// LS Electric XG5000 project: EV_s3
// PLC LSPLC
// module base 0 slot 0: 입출력 모듈:XBC-DR32H (DC 24V 입력, 릴레이 출력 32점)
// module base 0 slot 1: 입력 모듈:XBE-DC16A/B (DC24V 입력, 16점 / DC12/24V 입력, 16점)
// module base 0 slot 2: FEnet:XBL-EMTA (Ethernet 통신 모듈, 전기 Master)
// task INIT: Kind=1 Priority=2

PROGRAM VFD_PARAM (task: 스캔 프로그램)

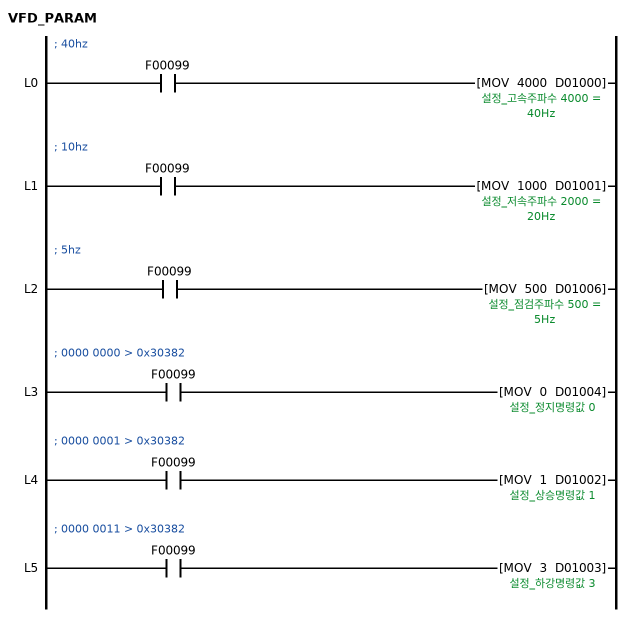
; L0
LOAD      F00099
MOV       4000 D01000	// 설정_고속주파수 4000 = 40Hz
// output comment: 40hz
; L1
LOAD      F00099
MOV       1000 D01001	// 설정_저속주파수 2000 = 20Hz
// output comment: 10hz
; L2
LOAD      F00099
MOV       500 D01006	// 설정_점검주파수 500 = 5Hz
// output comment: 5hz
; L3
LOAD      F00099
MOV       0 D01004	// 설정_정지명령값 0
// output comment: 0000 0000 > 0x30382
; L4
LOAD      F00099
MOV       1 D01002	// 설정_상승명령값 1
// output comment: 0000 0001 > 0x30382
; L5
LOAD      F00099
MOV       3 D01003	// 설정_하강명령값 3
// output comment: 0000 0011 > 0x30382

PROGRAM P00_P_MIRROR (task: 스캔 프로그램)

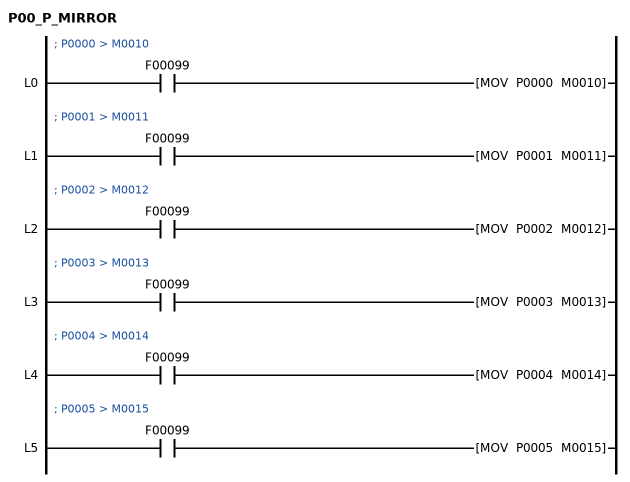
; L0
LOAD      F00099
MOV       P0000 M0010
// output comment: P0000 > M0010
; L1
LOAD      F00099
MOV       P0001 M0011
// output comment: P0001 > M0011
; L2
LOAD      F00099
MOV       P0002 M0012
// output comment: P0002 > M0012
; L3
LOAD      F00099
MOV       P0003 M0013
// output comment: P0003 > M0013
; L4
LOAD      F00099
MOV       P0004 M0014
// output comment: P0004 > M0014
; L5
LOAD      F00099
MOV       P0005 M0015
// output comment: P0005 > M0015

PROGRAM P01_POSITION (task: 스캔 프로그램)

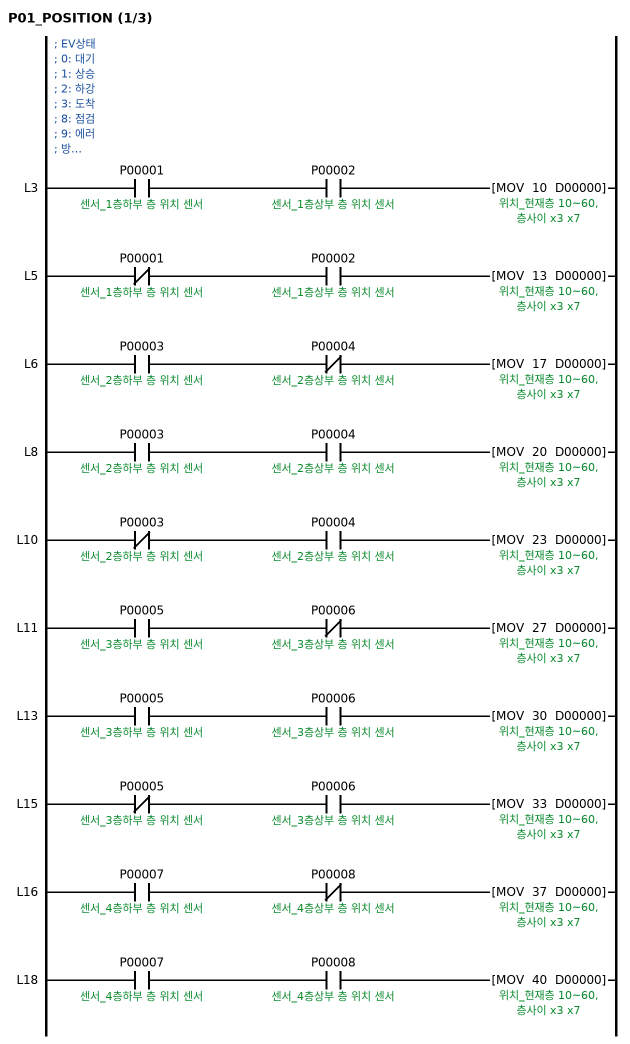
// EV상태
// 0: 대기
// 1: 상승
// 2: 하강
// 3: 도착
// 8: 점검
// 9: 에러
// 방향
// 0: 대기
// 1: 상승
// 2: 하강
// 센서로 인한 현재 위치
; L3
LOAD      P00001	// 센서_1층하부 층 위치 센서
AND       P00002	// 센서_1층상부 층 위치 센서
MOV       10 D00000	// 위치_현재층 10~60, 층사이 x3 x7
; L5
LOAD NOT  P00001	// 센서_1층하부 층 위치 센서
AND       P00002	// 센서_1층상부 층 위치 센서
MOV       13 D00000	// 위치_현재층 10~60, 층사이 x3 x7
; L6
LOAD      P00003	// 센서_2층하부 층 위치 센서
AND NOT   P00004	// 센서_2층상부 층 위치 센서
MOV       17 D00000	// 위치_현재층 10~60, 층사이 x3 x7
; L8
LOAD      P00003	// 센서_2층하부 층 위치 센서
AND       P00004	// 센서_2층상부 층 위치 센서
MOV       20 D00000	// 위치_현재층 10~60, 층사이 x3 x7
; L10
LOAD NOT  P00003	// 센서_2층하부 층 위치 센서
AND       P00004	// 센서_2층상부 층 위치 센서
MOV       23 D00000	// 위치_현재층 10~60, 층사이 x3 x7
; L11
LOAD      P00005	// 센서_3층하부 층 위치 센서
AND NOT   P00006	// 센서_3층상부 층 위치 센서
MOV       27 D00000	// 위치_현재층 10~60, 층사이 x3 x7
; L13
LOAD      P00005	// 센서_3층하부 층 위치 센서
AND       P00006	// 센서_3층상부 층 위치 센서
MOV       30 D00000	// 위치_현재층 10~60, 층사이 x3 x7
; L15
LOAD NOT  P00005	// 센서_3층하부 층 위치 센서
AND       P00006	// 센서_3층상부 층 위치 센서
MOV       33 D00000	// 위치_현재층 10~60, 층사이 x3 x7
; L16
LOAD      P00007	// 센서_4층하부 층 위치 센서
AND NOT   P00008	// 센서_4층상부 층 위치 센서
MOV       37 D00000	// 위치_현재층 10~60, 층사이 x3 x7
; L18
LOAD      P00007	// 센서_4층하부 층 위치 센서
AND       P00008	// 센서_4층상부 층 위치 센서
MOV       40 D00000	// 위치_현재층 10~60, 층사이 x3 x7

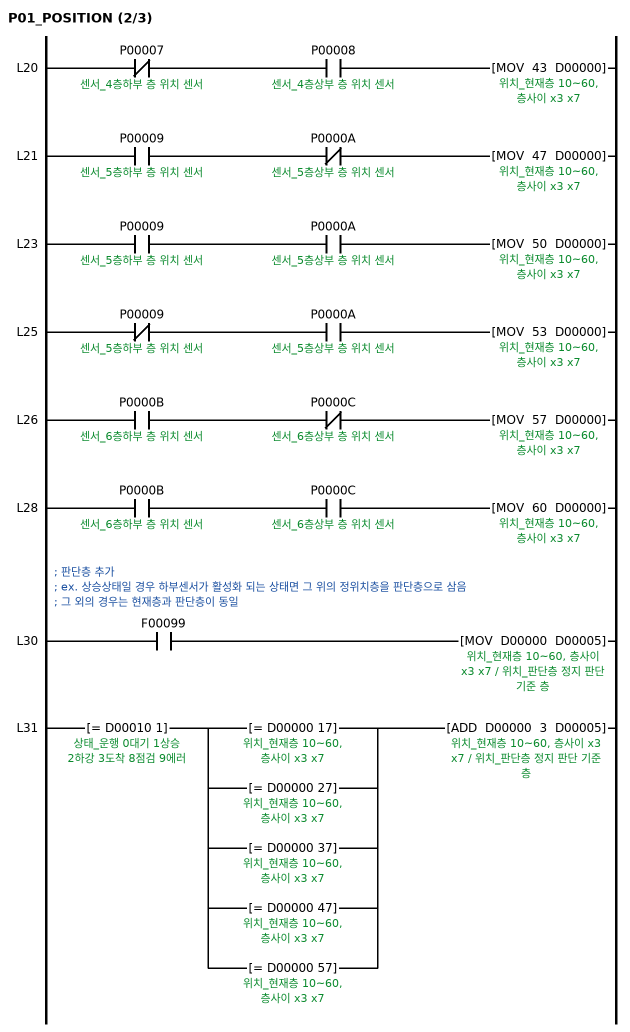
; L20
LOAD NOT  P00007	// 센서_4층하부 층 위치 센서
AND       P00008	// 센서_4층상부 층 위치 센서
MOV       43 D00000	// 위치_현재층 10~60, 층사이 x3 x7
; L21
LOAD      P00009	// 센서_5층하부 층 위치 센서
AND NOT   P0000A	// 센서_5층상부 층 위치 센서
MOV       47 D00000	// 위치_현재층 10~60, 층사이 x3 x7
; L23
LOAD      P00009	// 센서_5층하부 층 위치 센서
AND       P0000A	// 센서_5층상부 층 위치 센서
MOV       50 D00000	// 위치_현재층 10~60, 층사이 x3 x7
; L25
LOAD NOT  P00009	// 센서_5층하부 층 위치 센서
AND       P0000A	// 센서_5층상부 층 위치 센서
MOV       53 D00000	// 위치_현재층 10~60, 층사이 x3 x7
; L26
LOAD      P0000B	// 센서_6층하부 층 위치 센서
AND NOT   P0000C	// 센서_6층상부 층 위치 센서
MOV       57 D00000	// 위치_현재층 10~60, 층사이 x3 x7
; L28
LOAD      P0000B	// 센서_6층하부 층 위치 센서
AND       P0000C	// 센서_6층상부 층 위치 센서
MOV       60 D00000	// 위치_현재층 10~60, 층사이 x3 x7
// 판단층 추가
// ex. 상승상태일 경우 하부센서가 활성화 되는 상태면 그 위의 정위치층을 판단층으로 삼음
// 그 외의 경우는 현재층과 판단층이 동일
; L30
LOAD      F00099
MOV       D00000 D00005	// 위치_현재층 10~60, 층사이 x3 x7 / 위치_판단층 정지 판단 기준 층
; L31
LOAD=     D00010 1	// 상태_운행 0대기 1상승 2하강 3도착 8점검 9에러
LOAD=     D00000 17	// 위치_현재층 10~60, 층사이 x3 x7
OR=       D00000 27	// 위치_현재층 10~60, 층사이 x3 x7
OR=       D00000 37	// 위치_현재층 10~60, 층사이 x3 x7
OR=       D00000 47	// 위치_현재층 10~60, 층사이 x3 x7
OR=       D00000 57	// 위치_현재층 10~60, 층사이 x3 x7
AND LOAD
ADD       D00000 3 D00005	// 위치_현재층 10~60, 층사이 x3 x7 / 위치_판단층 정지 판단 기준 층

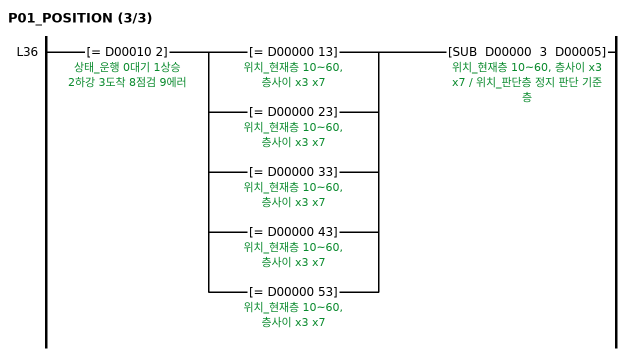
; L36
LOAD=     D00010 2	// 상태_운행 0대기 1상승 2하강 3도착 8점검 9에러
LOAD=     D00000 13	// 위치_현재층 10~60, 층사이 x3 x7
OR=       D00000 23	// 위치_현재층 10~60, 층사이 x3 x7
OR=       D00000 33	// 위치_현재층 10~60, 층사이 x3 x7
OR=       D00000 43	// 위치_현재층 10~60, 층사이 x3 x7
OR=       D00000 53	// 위치_현재층 10~60, 층사이 x3 x7
AND LOAD
SUB       D00000 3 D00005	// 위치_현재층 10~60, 층사이 x3 x7 / 위치_판단층 정지 판단 기준 층

PROGRAM P02_REQUEST (task: 스캔 프로그램)

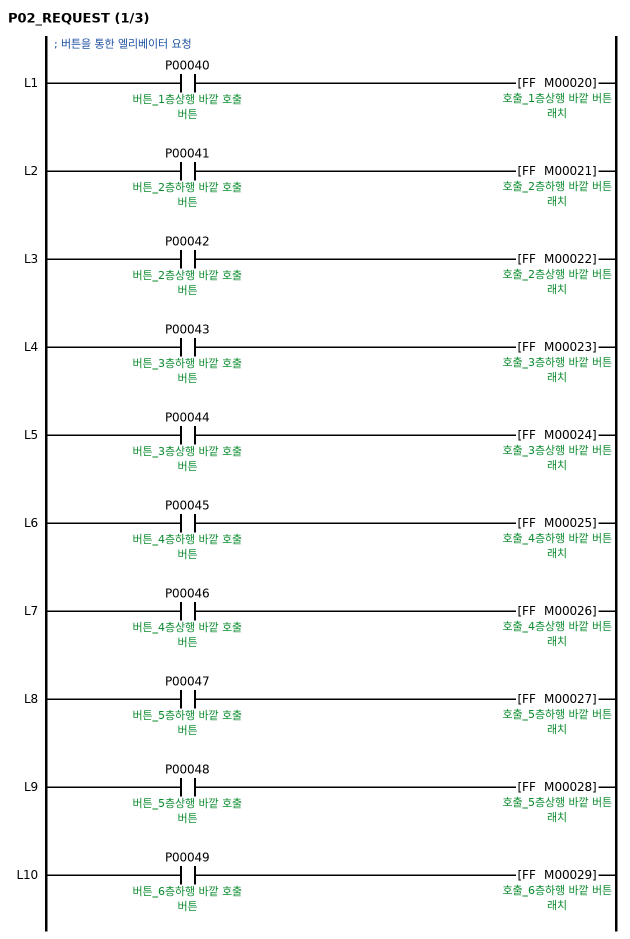
// 버튼을 통한 엘리베이터 요청
; L1
LOAD      P00040	// 버튼_1층상행 바깥 호출 버튼
FF        M00020	// 호출_1층상행 바깥 버튼 래치
; L2
LOAD      P00041	// 버튼_2층하행 바깥 호출 버튼
FF        M00021	// 호출_2층하행 바깥 버튼 래치
; L3
LOAD      P00042	// 버튼_2층상행 바깥 호출 버튼
FF        M00022	// 호출_2층상행 바깥 버튼 래치
; L4
LOAD      P00043	// 버튼_3층하행 바깥 호출 버튼
FF        M00023	// 호출_3층하행 바깥 버튼 래치
; L5
LOAD      P00044	// 버튼_3층상행 바깥 호출 버튼
FF        M00024	// 호출_3층상행 바깥 버튼 래치
; L6
LOAD      P00045	// 버튼_4층하행 바깥 호출 버튼
FF        M00025	// 호출_4층하행 바깥 버튼 래치
; L7
LOAD      P00046	// 버튼_4층상행 바깥 호출 버튼
FF        M00026	// 호출_4층상행 바깥 버튼 래치
; L8
LOAD      P00047	// 버튼_5층하행 바깥 호출 버튼
FF        M00027	// 호출_5층하행 바깥 버튼 래치
; L9
LOAD      P00048	// 버튼_5층상행 바깥 호출 버튼
FF        M00028	// 호출_5층상행 바깥 버튼 래치
; L10
LOAD      P00049	// 버튼_6층하행 바깥 호출 버튼
FF        M00029	// 호출_6층하행 바깥 버튼 래치

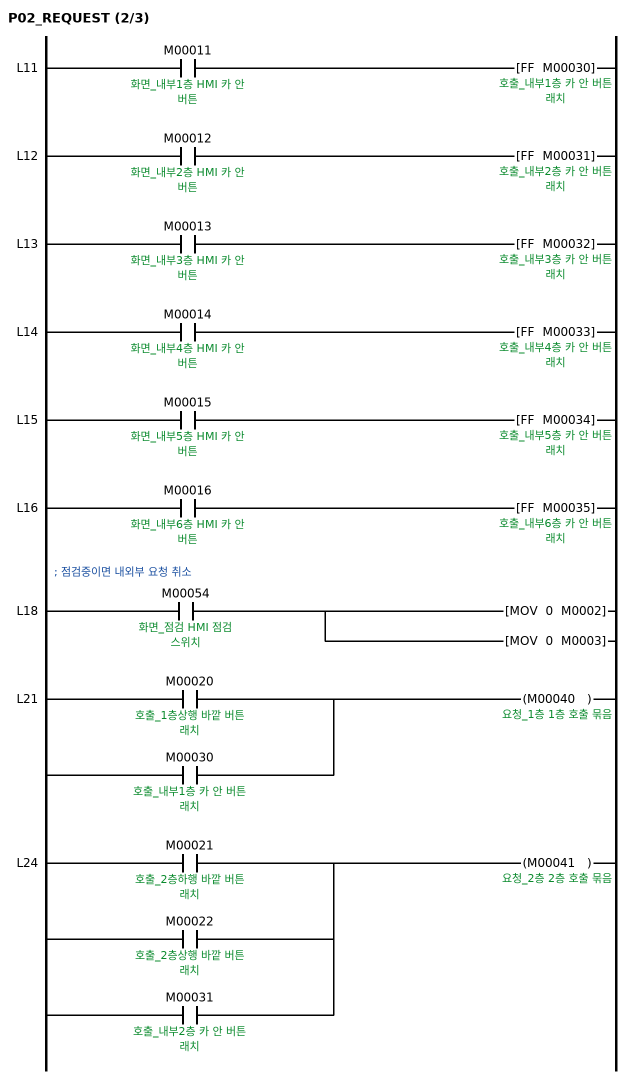
; L11
LOAD      M00011	// 화면_내부1층 HMI 카 안 버튼
FF        M00030	// 호출_내부1층 카 안 버튼 래치
; L12
LOAD      M00012	// 화면_내부2층 HMI 카 안 버튼
FF        M00031	// 호출_내부2층 카 안 버튼 래치
; L13
LOAD      M00013	// 화면_내부3층 HMI 카 안 버튼
FF        M00032	// 호출_내부3층 카 안 버튼 래치
; L14
LOAD      M00014	// 화면_내부4층 HMI 카 안 버튼
FF        M00033	// 호출_내부4층 카 안 버튼 래치
; L15
LOAD      M00015	// 화면_내부5층 HMI 카 안 버튼
FF        M00034	// 호출_내부5층 카 안 버튼 래치
; L16
LOAD      M00016	// 화면_내부6층 HMI 카 안 버튼
FF        M00035	// 호출_내부6층 카 안 버튼 래치
; L18
LOAD      M00054	// 화면_점검 HMI 점검 스위치
MOV       0 M0002
MOV       0 M0003
// output comment: 점검중이면 내외부 요청 취소
; L21
LOAD      M00020	// 호출_1층상행 바깥 버튼 래치
OR        M00030	// 호출_내부1층 카 안 버튼 래치
OUT       M00040	// 요청_1층 1층 호출 묶음
; L24
LOAD      M00021	// 호출_2층하행 바깥 버튼 래치
OR        M00022	// 호출_2층상행 바깥 버튼 래치
OR        M00031	// 호출_내부2층 카 안 버튼 래치
OUT       M00041	// 요청_2층 2층 호출 묶음

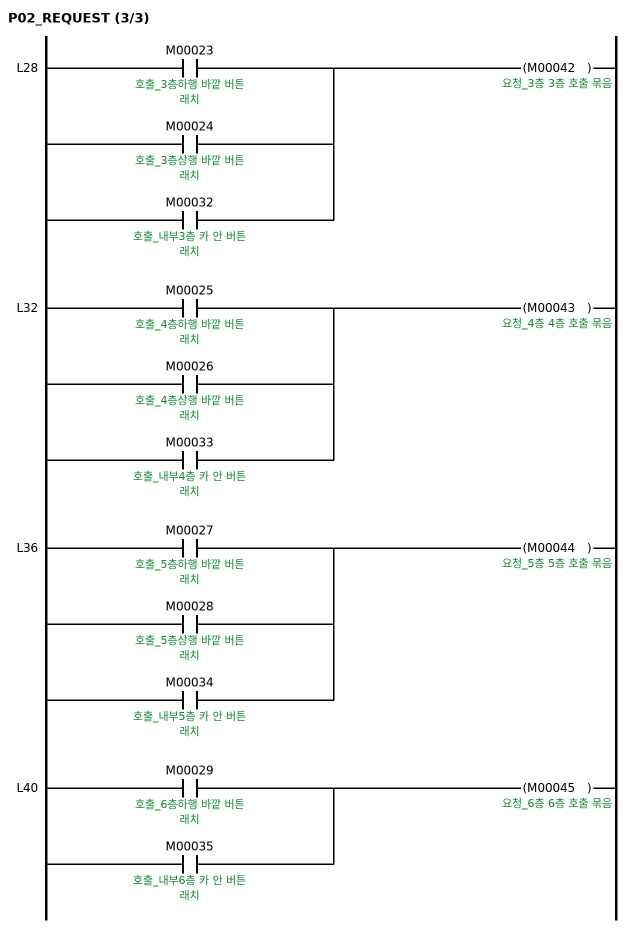
; L28
LOAD      M00023	// 호출_3층하행 바깥 버튼 래치
OR        M00024	// 호출_3층상행 바깥 버튼 래치
OR        M00032	// 호출_내부3층 카 안 버튼 래치
OUT       M00042	// 요청_3층 3층 호출 묶음
; L32
LOAD      M00025	// 호출_4층하행 바깥 버튼 래치
OR        M00026	// 호출_4층상행 바깥 버튼 래치
OR        M00033	// 호출_내부4층 카 안 버튼 래치
OUT       M00043	// 요청_4층 4층 호출 묶음
; L36
LOAD      M00027	// 호출_5층하행 바깥 버튼 래치
OR        M00028	// 호출_5층상행 바깥 버튼 래치
OR        M00034	// 호출_내부5층 카 안 버튼 래치
OUT       M00044	// 요청_5층 5층 호출 묶음
; L40
LOAD      M00029	// 호출_6층하행 바깥 버튼 래치
OR        M00035	// 호출_내부6층 카 안 버튼 래치
OUT       M00045	// 요청_6층 6층 호출 묶음

PROGRAM P03_JUDGE (task: 스캔 프로그램)

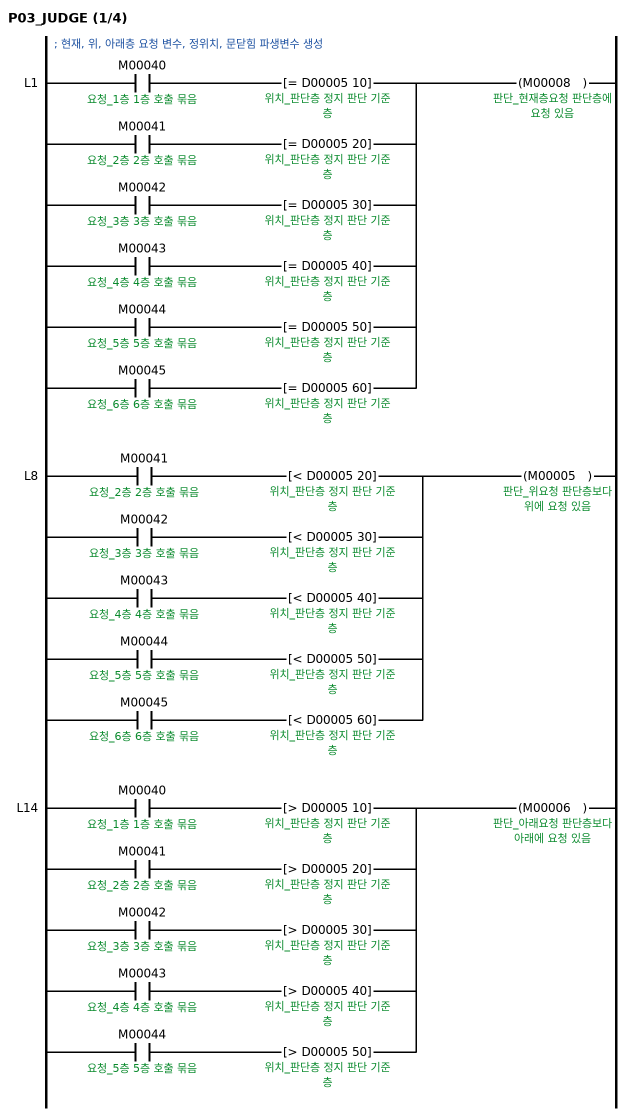
// 현재, 위, 아래층 요청 변수, 정위치, 문닫힘 파생변수 생성
; L1
LOAD      M00040	// 요청_1층 1층 호출 묶음
AND=      D00005 10	// 위치_판단층 정지 판단 기준 층
LOAD      M00041	// 요청_2층 2층 호출 묶음
AND=      D00005 20	// 위치_판단층 정지 판단 기준 층
OR LOAD
LOAD      M00042	// 요청_3층 3층 호출 묶음
AND=      D00005 30	// 위치_판단층 정지 판단 기준 층
OR LOAD
LOAD      M00043	// 요청_4층 4층 호출 묶음
AND=      D00005 40	// 위치_판단층 정지 판단 기준 층
OR LOAD
LOAD      M00044	// 요청_5층 5층 호출 묶음
AND=      D00005 50	// 위치_판단층 정지 판단 기준 층
OR LOAD
LOAD      M00045	// 요청_6층 6층 호출 묶음
AND=      D00005 60	// 위치_판단층 정지 판단 기준 층
OR LOAD
OUT       M00008	// 판단_현재층요청 판단층에 요청 있음
; L8
LOAD      M00041	// 요청_2층 2층 호출 묶음
AND<      D00005 20	// 위치_판단층 정지 판단 기준 층
LOAD      M00042	// 요청_3층 3층 호출 묶음
AND<      D00005 30	// 위치_판단층 정지 판단 기준 층
OR LOAD
LOAD      M00043	// 요청_4층 4층 호출 묶음
AND<      D00005 40	// 위치_판단층 정지 판단 기준 층
OR LOAD
LOAD      M00044	// 요청_5층 5층 호출 묶음
AND<      D00005 50	// 위치_판단층 정지 판단 기준 층
OR LOAD
LOAD      M00045	// 요청_6층 6층 호출 묶음
AND<      D00005 60	// 위치_판단층 정지 판단 기준 층
OR LOAD
OUT       M00005	// 판단_위요청 판단층보다 위에 요청 있음
; L14
LOAD      M00040	// 요청_1층 1층 호출 묶음
AND>      D00005 10	// 위치_판단층 정지 판단 기준 층
LOAD      M00041	// 요청_2층 2층 호출 묶음
AND>      D00005 20	// 위치_판단층 정지 판단 기준 층
OR LOAD
LOAD      M00042	// 요청_3층 3층 호출 묶음
AND>      D00005 30	// 위치_판단층 정지 판단 기준 층
OR LOAD
LOAD      M00043	// 요청_4층 4층 호출 묶음
AND>      D00005 40	// 위치_판단층 정지 판단 기준 층
OR LOAD
LOAD      M00044	// 요청_5층 5층 호출 묶음
AND>      D00005 50	// 위치_판단층 정지 판단 기준 층
OR LOAD
OUT       M00006	// 판단_아래요청 판단층보다 아래에 요청 있음

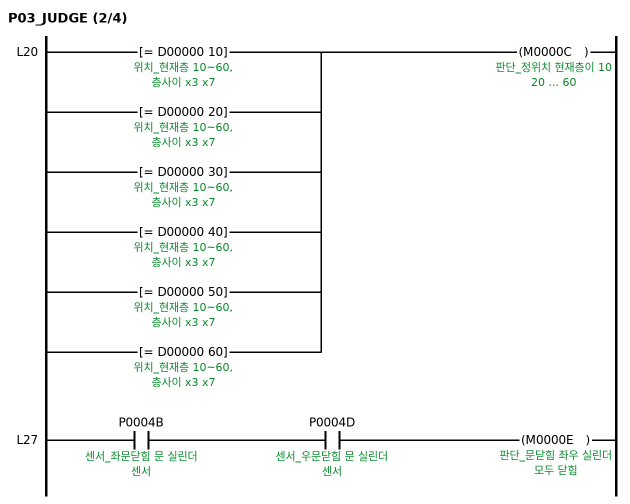
; L20
LOAD=     D00000 10	// 위치_현재층 10~60, 층사이 x3 x7
OR=       D00000 20	// 위치_현재층 10~60, 층사이 x3 x7
OR=       D00000 30	// 위치_현재층 10~60, 층사이 x3 x7
OR=       D00000 40	// 위치_현재층 10~60, 층사이 x3 x7
OR=       D00000 50	// 위치_현재층 10~60, 층사이 x3 x7
OR=       D00000 60	// 위치_현재층 10~60, 층사이 x3 x7
OUT       M0000C	// 판단_정위치 현재층이 10 20 ... 60
; L27
LOAD      P0004B	// 센서_좌문닫힘 문 실린더 센서
AND       P0004D	// 센서_우문닫힘 문 실린더 센서
OUT       M0000E	// 판단_문닫힘 좌우 실린더 모두 닫힘

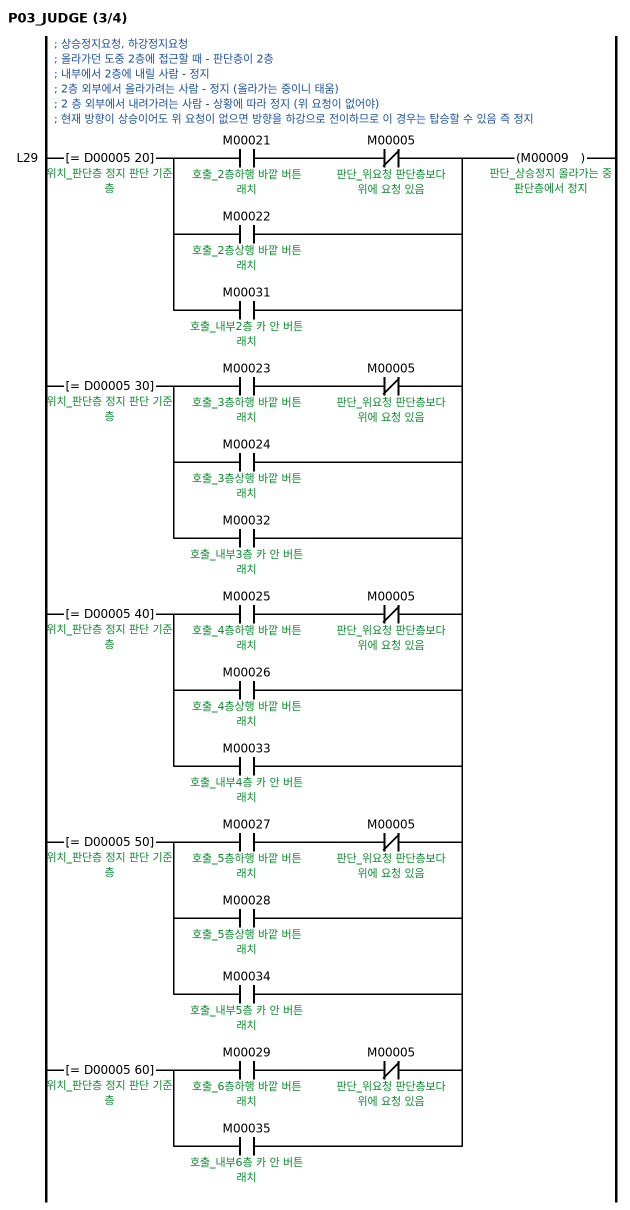
// 상승정지요청, 하강정지요청
; L29
LOAD=     D00005 20	// 위치_판단층 정지 판단 기준 층
LOAD      M00021	// 호출_2층하행 바깥 버튼 래치
AND NOT   M00005	// 판단_위요청 판단층보다 위에 요청 있음
OR        M00022	// 호출_2층상행 바깥 버튼 래치
OR        M00031	// 호출_내부2층 카 안 버튼 래치
AND LOAD
LOAD=     D00005 30	// 위치_판단층 정지 판단 기준 층
LOAD      M00023	// 호출_3층하행 바깥 버튼 래치
AND NOT   M00005	// 판단_위요청 판단층보다 위에 요청 있음
OR        M00024	// 호출_3층상행 바깥 버튼 래치
OR        M00032	// 호출_내부3층 카 안 버튼 래치
AND LOAD
OR LOAD
LOAD=     D00005 40	// 위치_판단층 정지 판단 기준 층
LOAD      M00025	// 호출_4층하행 바깥 버튼 래치
AND NOT   M00005	// 판단_위요청 판단층보다 위에 요청 있음
OR        M00026	// 호출_4층상행 바깥 버튼 래치
OR        M00033	// 호출_내부4층 카 안 버튼 래치
AND LOAD
OR LOAD
LOAD=     D00005 50	// 위치_판단층 정지 판단 기준 층
LOAD      M00027	// 호출_5층하행 바깥 버튼 래치
AND NOT   M00005	// 판단_위요청 판단층보다 위에 요청 있음
OR        M00028	// 호출_5층상행 바깥 버튼 래치
OR        M00034	// 호출_내부5층 카 안 버튼 래치
AND LOAD
OR LOAD
LOAD=     D00005 60	// 위치_판단층 정지 판단 기준 층
LOAD      M00029	// 호출_6층하행 바깥 버튼 래치
AND NOT   M00005	// 판단_위요청 판단층보다 위에 요청 있음
OR        M00035	// 호출_내부6층 카 안 버튼 래치
AND LOAD
OR LOAD
OUT       M00009	// 판단_상승정지 올라가는 중 판단층에서 정지
// output comment: 올라가던 도중 2층에 접근할 때 - 판단층이 2층 내부에서 2층에 내릴 사람 - 정지 2층 외부에서 올라가려는 사람 - 정지 (올라가는 중이니 태움) 2 층 외부에서 내려가려는 사람 - 상황에 따라 정지 (위 요청이 없어야) 현재 방향이 상승이어도 위 요청이 없으면 방향을 하강으로 전이하므로 이 경우는 탑승할 수 있음 즉 정지

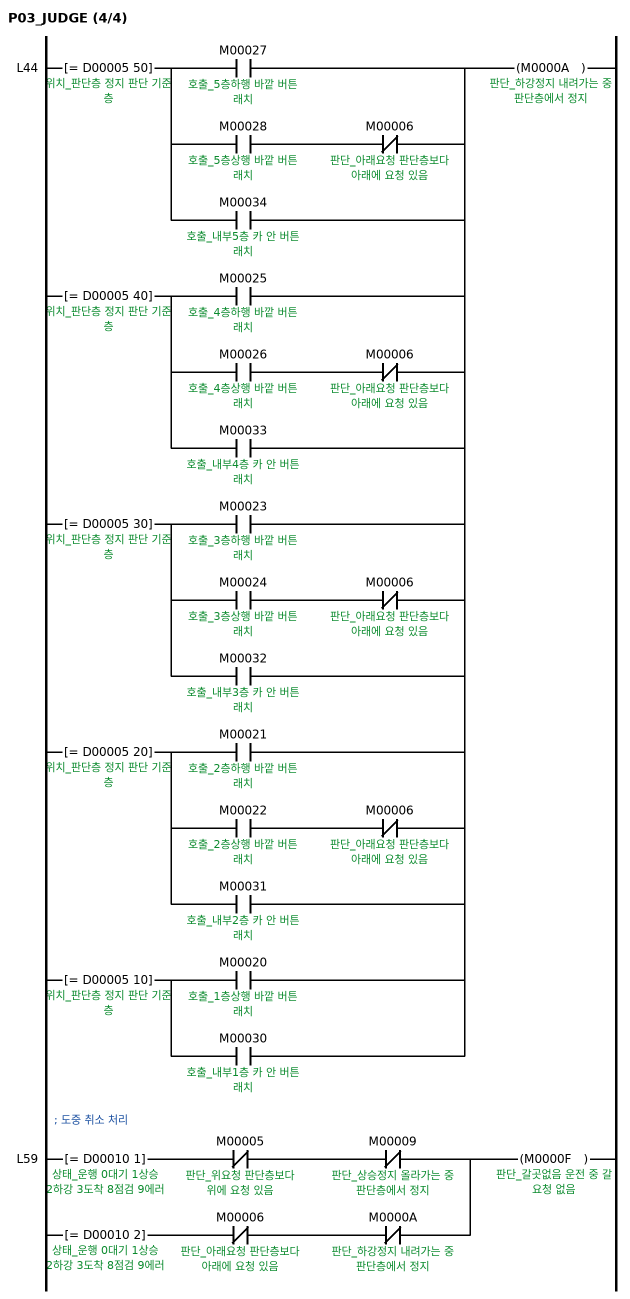
; L44
LOAD=     D00005 50	// 위치_판단층 정지 판단 기준 층
LOAD      M00027	// 호출_5층하행 바깥 버튼 래치
LOAD      M00028	// 호출_5층상행 바깥 버튼 래치
AND NOT   M00006	// 판단_아래요청 판단층보다 아래에 요청 있음
OR LOAD
OR        M00034	// 호출_내부5층 카 안 버튼 래치
AND LOAD
LOAD=     D00005 40	// 위치_판단층 정지 판단 기준 층
LOAD      M00025	// 호출_4층하행 바깥 버튼 래치
LOAD      M00026	// 호출_4층상행 바깥 버튼 래치
AND NOT   M00006	// 판단_아래요청 판단층보다 아래에 요청 있음
OR LOAD
OR        M00033	// 호출_내부4층 카 안 버튼 래치
AND LOAD
OR LOAD
LOAD=     D00005 30	// 위치_판단층 정지 판단 기준 층
LOAD      M00023	// 호출_3층하행 바깥 버튼 래치
LOAD      M00024	// 호출_3층상행 바깥 버튼 래치
AND NOT   M00006	// 판단_아래요청 판단층보다 아래에 요청 있음
OR LOAD
OR        M00032	// 호출_내부3층 카 안 버튼 래치
AND LOAD
OR LOAD
LOAD=     D00005 20	// 위치_판단층 정지 판단 기준 층
LOAD      M00021	// 호출_2층하행 바깥 버튼 래치
LOAD      M00022	// 호출_2층상행 바깥 버튼 래치
AND NOT   M00006	// 판단_아래요청 판단층보다 아래에 요청 있음
OR LOAD
OR        M00031	// 호출_내부2층 카 안 버튼 래치
AND LOAD
OR LOAD
LOAD=     D00005 10	// 위치_판단층 정지 판단 기준 층
LOAD      M00020	// 호출_1층상행 바깥 버튼 래치
OR        M00030	// 호출_내부1층 카 안 버튼 래치
AND LOAD
OR LOAD
OUT       M0000A	// 판단_하강정지 내려가는 중 판단층에서 정지
// 도중 취소 처리
; L59
LOAD=     D00010 1	// 상태_운행 0대기 1상승 2하강 3도착 8점검 9에러
AND NOT   M00005	// 판단_위요청 판단층보다 위에 요청 있음
AND NOT   M00009	// 판단_상승정지 올라가는 중 판단층에서 정지
LOAD=     D00010 2	// 상태_운행 0대기 1상승 2하강 3도착 8점검 9에러
AND NOT   M00006	// 판단_아래요청 판단층보다 아래에 요청 있음
AND NOT   M0000A	// 판단_하강정지 내려가는 중 판단층에서 정지
OR LOAD
OUT       M0000F	// 판단_갈곳없음 운전 중 갈 요청 없음

PROGRAM P04_TRANSITION (task: 스캔 프로그램)

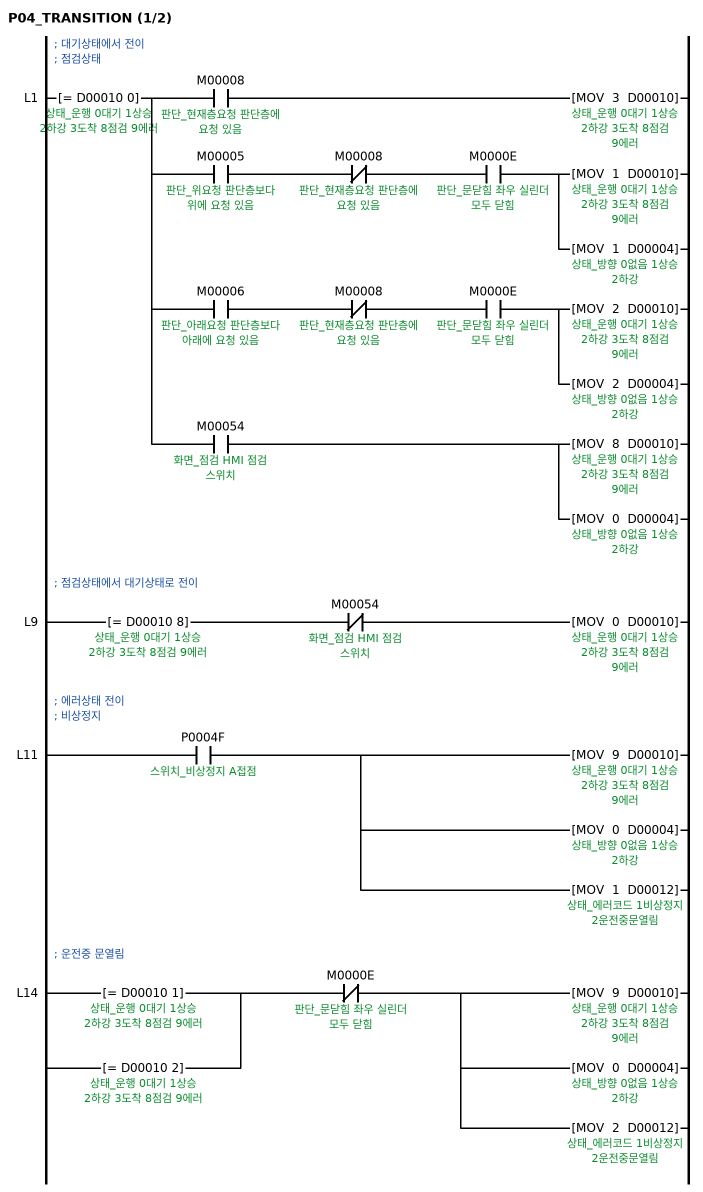
// 대기상태에서 전이
; L1
LOAD=     D00010 0	// 상태_운행 0대기 1상승 2하강 3도착 8점검 9에러
MPUSH
AND       M00008	// 판단_현재층요청 판단층에 요청 있음
MOV       3 D00010	// 상태_운행 0대기 1상승 2하강 3도착 8점검 9에러
MLOAD
AND       M00005	// 판단_위요청 판단층보다 위에 요청 있음
AND NOT   M00008	// 판단_현재층요청 판단층에 요청 있음
AND       M0000E	// 판단_문닫힘 좌우 실린더 모두 닫힘
MOV       1 D00010	// 상태_운행 0대기 1상승 2하강 3도착 8점검 9에러
MOV       1 D00004	// 상태_방향 0없음 1상승 2하강
MLOAD
AND       M00006	// 판단_아래요청 판단층보다 아래에 요청 있음
AND NOT   M00008	// 판단_현재층요청 판단층에 요청 있음
AND       M0000E	// 판단_문닫힘 좌우 실린더 모두 닫힘
MOV       2 D00010	// 상태_운행 0대기 1상승 2하강 3도착 8점검 9에러
MOV       2 D00004	// 상태_방향 0없음 1상승 2하강
MPOP
AND       M00054	// 화면_점검 HMI 점검 스위치
MOV       8 D00010	// 상태_운행 0대기 1상승 2하강 3도착 8점검 9에러
MOV       0 D00004	// 상태_방향 0없음 1상승 2하강
// output comment: 점검상태
// 점검상태에서 대기상태로 전이
; L9
LOAD=     D00010 8	// 상태_운행 0대기 1상승 2하강 3도착 8점검 9에러
AND NOT   M00054	// 화면_점검 HMI 점검 스위치
MOV       0 D00010	// 상태_운행 0대기 1상승 2하강 3도착 8점검 9에러
// 에러상태 전이
; L11
LOAD      P0004F	// 스위치_비상정지 A접점
MOV       9 D00010	// 상태_운행 0대기 1상승 2하강 3도착 8점검 9에러
MOV       0 D00004	// 상태_방향 0없음 1상승 2하강
MOV       1 D00012	// 상태_에러코드 1비상정지 2운전중문열림
// output comment: 비상정지
; L14
LOAD=     D00010 1	// 상태_운행 0대기 1상승 2하강 3도착 8점검 9에러
OR=       D00010 2	// 상태_운행 0대기 1상승 2하강 3도착 8점검 9에러
AND NOT   M0000E	// 판단_문닫힘 좌우 실린더 모두 닫힘
MOV       9 D00010	// 상태_운행 0대기 1상승 2하강 3도착 8점검 9에러
MOV       0 D00004	// 상태_방향 0없음 1상승 2하강
MOV       2 D00012	// 상태_에러코드 1비상정지 2운전중문열림
// output comment: 운전중 문열림

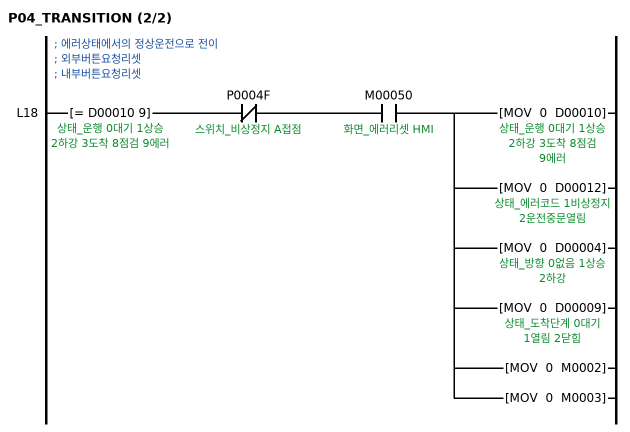
// 에러상태에서의 정상운전으로 전이
; L18
LOAD=     D00010 9	// 상태_운행 0대기 1상승 2하강 3도착 8점검 9에러
AND NOT   P0004F	// 스위치_비상정지 A접점
AND       M00050	// 화면_에러리셋 HMI
MOV       0 D00010	// 상태_운행 0대기 1상승 2하강 3도착 8점검 9에러
MOV       0 D00012	// 상태_에러코드 1비상정지 2운전중문열림
MOV       0 D00004	// 상태_방향 0없음 1상승 2하강
MOV       0 D00009	// 상태_도착단계 0대기 1열림 2닫힘
MOV       0 M0002
MOV       0 M0003
// output comment: 외부버튼요청리셋
// output comment: 내부버튼요청리셋

PROGRAM P05_DRIVE (task: 스캔 프로그램)

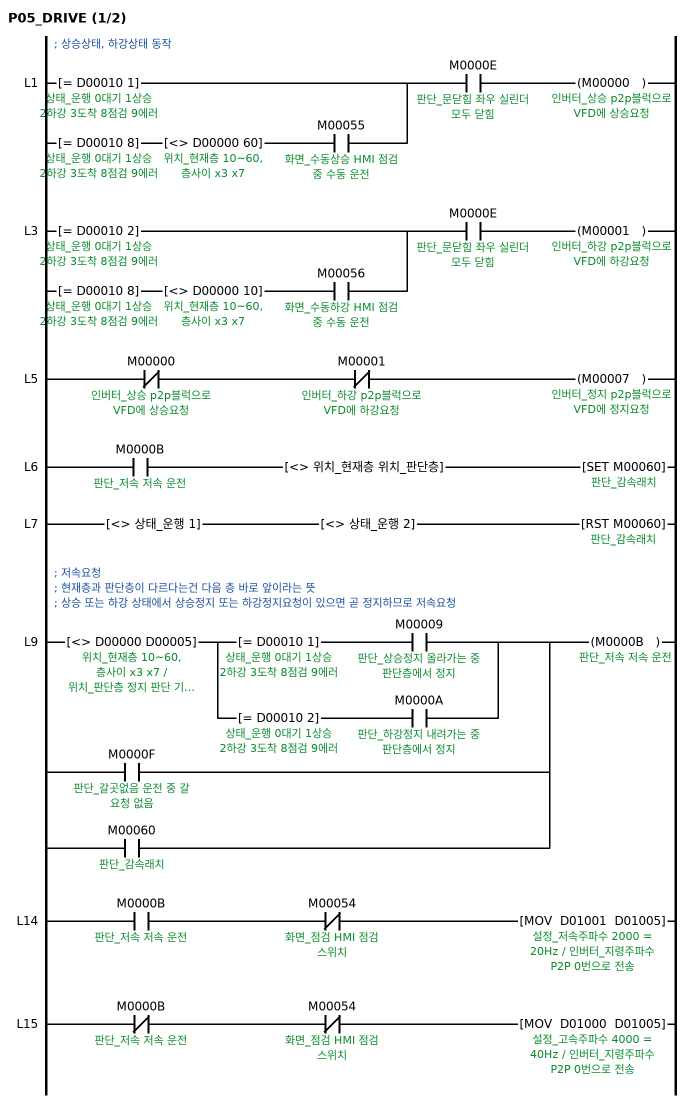
// 상승상태, 하강상태 동작
; L1
LOAD=     D00010 1	// 상태_운행 0대기 1상승 2하강 3도착 8점검 9에러
LOAD=     D00010 8	// 상태_운행 0대기 1상승 2하강 3도착 8점검 9에러
AND<>     D00000 60	// 위치_현재층 10~60, 층사이 x3 x7
AND       M00055	// 화면_수동상승 HMI 점검 중 수동 운전
OR LOAD
AND       M0000E	// 판단_문닫힘 좌우 실린더 모두 닫힘
OUT       M00000	// 인버터_상승 p2p블럭으로 VFD에 상승요청
; L3
LOAD=     D00010 2	// 상태_운행 0대기 1상승 2하강 3도착 8점검 9에러
LOAD=     D00010 8	// 상태_운행 0대기 1상승 2하강 3도착 8점검 9에러
AND<>     D00000 10	// 위치_현재층 10~60, 층사이 x3 x7
AND       M00056	// 화면_수동하강 HMI 점검 중 수동 운전
OR LOAD
AND       M0000E	// 판단_문닫힘 좌우 실린더 모두 닫힘
OUT       M00001	// 인버터_하강 p2p블럭으로 VFD에 하강요청
; L5
LOAD NOT  M00000	// 인버터_상승 p2p블럭으로 VFD에 상승요청
AND NOT   M00001	// 인버터_하강 p2p블럭으로 VFD에 하강요청
OUT       M00007	// 인버터_정지 p2p블럭으로 VFD에 정지요청
; L6
LOAD      M0000B	// 판단_저속 저속 운전
AND<>     위치_현재층 위치_판단층
SET       M00060	// 판단_감속래치
; L7
LOAD<>    상태_운행 1
AND<>     상태_운행 2
RST       M00060	// 판단_감속래치
// 저속요청
// 현재층과 판단층이 다르다는건 다음 층 바로 앞이라는 뜻 
// 상승 또는 하강 상태에서 상승정지 또는 하강정지요청이 있으면 곧 정지하므로 저속요청
; L9
LOAD<>    D00000 D00005	// 위치_현재층 10~60, 층사이 x3 x7 / 위치_판단층 정지 판단 기준 층
LOAD=     D00010 1	// 상태_운행 0대기 1상승 2하강 3도착 8점검 9에러
AND       M00009	// 판단_상승정지 올라가는 중 판단층에서 정지
LOAD=     D00010 2	// 상태_운행 0대기 1상승 2하강 3도착 8점검 9에러
AND       M0000A	// 판단_하강정지 내려가는 중 판단층에서 정지
OR LOAD
AND LOAD
OR        M0000F	// 판단_갈곳없음 운전 중 갈 요청 없음
OR        M00060	// 판단_감속래치
OUT       M0000B	// 판단_저속 저속 운전
; L14
LOAD      M0000B	// 판단_저속 저속 운전
AND NOT   M00054	// 화면_점검 HMI 점검 스위치
MOV       D01001 D01005	// 설정_저속주파수 2000 = 20Hz / 인버터_지령주파수 P2P 0번으로 전송
; L15
LOAD NOT  M0000B	// 판단_저속 저속 운전
AND NOT   M00054	// 화면_점검 HMI 점검 스위치
MOV       D01000 D01005	// 설정_고속주파수 4000 = 40Hz / 인버터_지령주파수 P2P 0번으로 전송

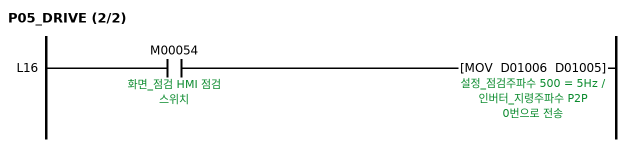
; L16
LOAD      M00054	// 화면_점검 HMI 점검 스위치
MOV       D01006 D01005	// 설정_점검주파수 500 = 5Hz / 인버터_지령주파수 P2P 0번으로 전송

PROGRAM P06_ARRIVE (task: 스캔 프로그램)

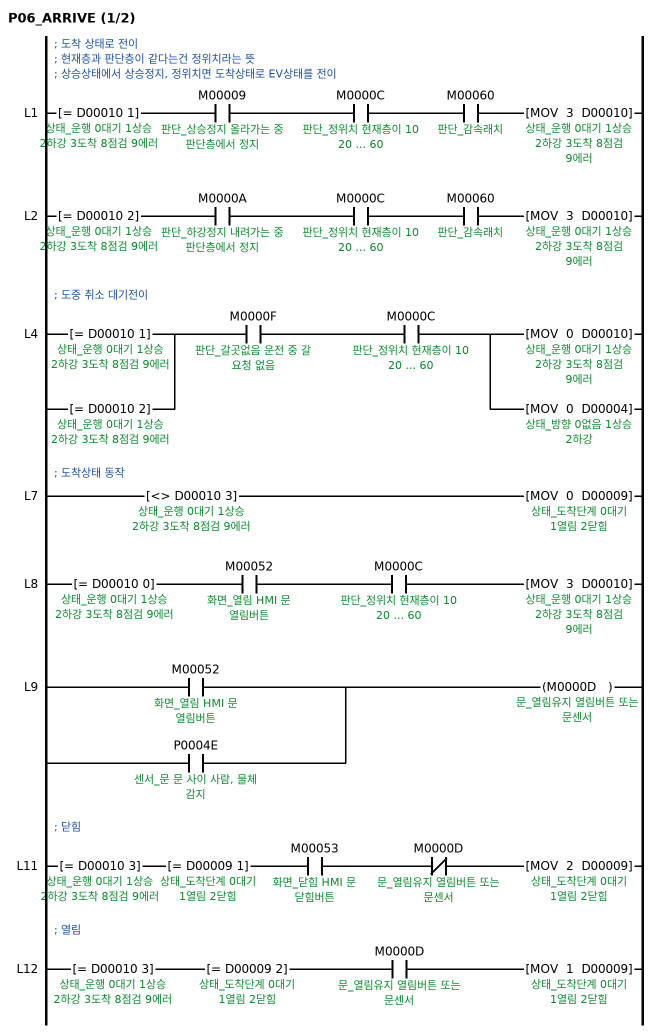
// 도착 상태로 전이
// 현재층과 판단층이 같다는건 정위치라는 뜻
// 상승상태에서 상승정지, 정위치면 도착상태로 EV상태를 전이
; L1
LOAD=     D00010 1	// 상태_운행 0대기 1상승 2하강 3도착 8점검 9에러
AND       M00009	// 판단_상승정지 올라가는 중 판단층에서 정지
AND       M0000C	// 판단_정위치 현재층이 10 20 ... 60
AND       M00060	// 판단_감속래치
MOV       3 D00010	// 상태_운행 0대기 1상승 2하강 3도착 8점검 9에러
; L2
LOAD=     D00010 2	// 상태_운행 0대기 1상승 2하강 3도착 8점검 9에러
AND       M0000A	// 판단_하강정지 내려가는 중 판단층에서 정지
AND       M0000C	// 판단_정위치 현재층이 10 20 ... 60
AND       M00060	// 판단_감속래치
MOV       3 D00010	// 상태_운행 0대기 1상승 2하강 3도착 8점검 9에러
// 도중 취소 대기전이
; L4
LOAD=     D00010 1	// 상태_운행 0대기 1상승 2하강 3도착 8점검 9에러
OR=       D00010 2	// 상태_운행 0대기 1상승 2하강 3도착 8점검 9에러
AND       M0000F	// 판단_갈곳없음 운전 중 갈 요청 없음
AND       M0000C	// 판단_정위치 현재층이 10 20 ... 60
MOV       0 D00010	// 상태_운행 0대기 1상승 2하강 3도착 8점검 9에러
MOV       0 D00004	// 상태_방향 0없음 1상승 2하강
// 도착상태 동작
; L7
LOAD<>    D00010 3	// 상태_운행 0대기 1상승 2하강 3도착 8점검 9에러
MOV       0 D00009	// 상태_도착단계 0대기 1열림 2닫힘
; L8
LOAD=     D00010 0	// 상태_운행 0대기 1상승 2하강 3도착 8점검 9에러
AND       M00052	// 화면_열림 HMI 문 열림버튼
AND       M0000C	// 판단_정위치 현재층이 10 20 ... 60
MOV       3 D00010	// 상태_운행 0대기 1상승 2하강 3도착 8점검 9에러
; L9
LOAD      M00052	// 화면_열림 HMI 문 열림버튼
OR        P0004E	// 센서_문 문 사이 사람, 물체 감지
OUT       M0000D	// 문_열림유지 열림버튼 또는 문센서
; L11
LOAD=     D00010 3	// 상태_운행 0대기 1상승 2하강 3도착 8점검 9에러
AND=      D00009 1	// 상태_도착단계 0대기 1열림 2닫힘
AND       M00053	// 화면_닫힘 HMI 문 닫힘버튼
AND NOT   M0000D	// 문_열림유지 열림버튼 또는 문센서
MOV       2 D00009	// 상태_도착단계 0대기 1열림 2닫힘
// output comment: 닫힘
; L12
LOAD=     D00010 3	// 상태_운행 0대기 1상승 2하강 3도착 8점검 9에러
AND=      D00009 2	// 상태_도착단계 0대기 1열림 2닫힘
AND       M0000D	// 문_열림유지 열림버튼 또는 문센서
MOV       1 D00009	// 상태_도착단계 0대기 1열림 2닫힘
// output comment: 열림

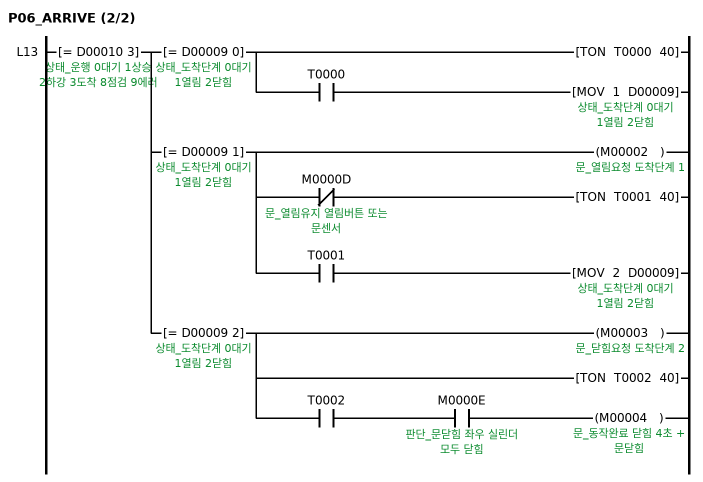
; L13
LOAD=     D00010 3	// 상태_운행 0대기 1상승 2하강 3도착 8점검 9에러
MPUSH
AND=      D00009 0	// 상태_도착단계 0대기 1열림 2닫힘
TON       T0000 40
AND       T0000
MOV       1 D00009	// 상태_도착단계 0대기 1열림 2닫힘
MLOAD
AND=      D00009 1	// 상태_도착단계 0대기 1열림 2닫힘
OUT       M00002	// 문_열림요청 도착단계 1
MPUSH
AND NOT   M0000D	// 문_열림유지 열림버튼 또는 문센서
TON       T0001 40
MPOP
AND       T0001
MOV       2 D00009	// 상태_도착단계 0대기 1열림 2닫힘
MPOP
AND=      D00009 2	// 상태_도착단계 0대기 1열림 2닫힘
OUT       M00003	// 문_닫힘요청 도착단계 2
TON       T0002 40
AND       T0002
AND       M0000E	// 판단_문닫힘 좌우 실린더 모두 닫힘
OUT       M00004	// 문_동작완료 닫힘 4초 + 문닫힘

PROGRAM P07_DISPATCH (task: 스캔 프로그램)

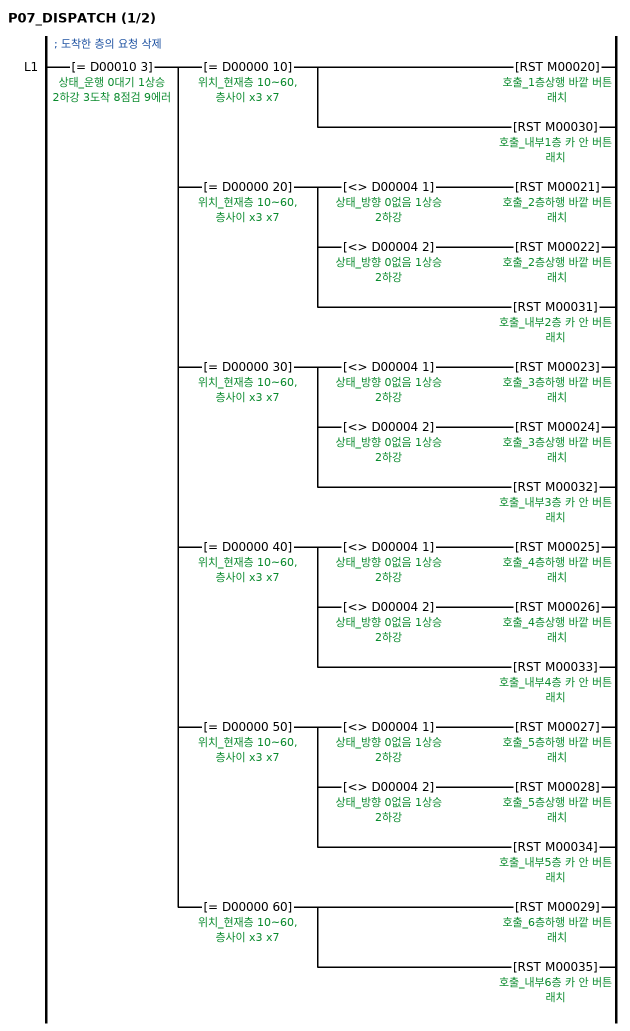
// 도착한 층의 요청 삭제
; L1
LOAD=     D00010 3	// 상태_운행 0대기 1상승 2하강 3도착 8점검 9에러
MPUSH
AND=      D00000 10	// 위치_현재층 10~60, 층사이 x3 x7
RST       M00020	// 호출_1층상행 바깥 버튼 래치
RST       M00030	// 호출_내부1층 카 안 버튼 래치
MLOAD
AND=      D00000 20	// 위치_현재층 10~60, 층사이 x3 x7
MPUSH
AND<>     D00004 1	// 상태_방향 0없음 1상승 2하강
RST       M00021	// 호출_2층하행 바깥 버튼 래치
MLOAD
AND<>     D00004 2	// 상태_방향 0없음 1상승 2하강
RST       M00022	// 호출_2층상행 바깥 버튼 래치
MPOP
RST       M00031	// 호출_내부2층 카 안 버튼 래치
MLOAD
AND=      D00000 30	// 위치_현재층 10~60, 층사이 x3 x7
MPUSH
AND<>     D00004 1	// 상태_방향 0없음 1상승 2하강
RST       M00023	// 호출_3층하행 바깥 버튼 래치
MLOAD
AND<>     D00004 2	// 상태_방향 0없음 1상승 2하강
RST       M00024	// 호출_3층상행 바깥 버튼 래치
MPOP
RST       M00032	// 호출_내부3층 카 안 버튼 래치
MLOAD
AND=      D00000 40	// 위치_현재층 10~60, 층사이 x3 x7
MPUSH
AND<>     D00004 1	// 상태_방향 0없음 1상승 2하강
RST       M00025	// 호출_4층하행 바깥 버튼 래치
MLOAD
AND<>     D00004 2	// 상태_방향 0없음 1상승 2하강
RST       M00026	// 호출_4층상행 바깥 버튼 래치
MPOP
RST       M00033	// 호출_내부4층 카 안 버튼 래치
MLOAD
AND=      D00000 50	// 위치_현재층 10~60, 층사이 x3 x7
MPUSH
AND<>     D00004 1	// 상태_방향 0없음 1상승 2하강
RST       M00027	// 호출_5층하행 바깥 버튼 래치
MLOAD
AND<>     D00004 2	// 상태_방향 0없음 1상승 2하강
RST       M00028	// 호출_5층상행 바깥 버튼 래치
MPOP
RST       M00034	// 호출_내부5층 카 안 버튼 래치
MPOP
AND=      D00000 60	// 위치_현재층 10~60, 층사이 x3 x7
RST       M00029	// 호출_6층하행 바깥 버튼 래치
RST       M00035	// 호출_내부6층 카 안 버튼 래치

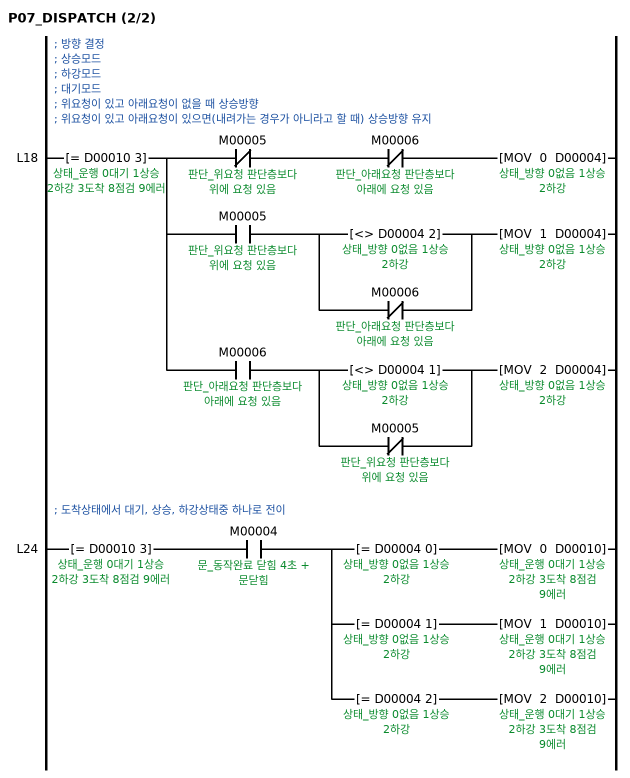
// 방향 결정
// 상승모드
// 하강모드
// 대기모드
; L18
LOAD=     D00010 3	// 상태_운행 0대기 1상승 2하강 3도착 8점검 9에러
MPUSH
AND NOT   M00005	// 판단_위요청 판단층보다 위에 요청 있음
AND NOT   M00006	// 판단_아래요청 판단층보다 아래에 요청 있음
MOV       0 D00004	// 상태_방향 0없음 1상승 2하강
MLOAD
AND       M00005	// 판단_위요청 판단층보다 위에 요청 있음
LOAD<>    D00004 2	// 상태_방향 0없음 1상승 2하강
OR NOT    M00006	// 판단_아래요청 판단층보다 아래에 요청 있음
AND LOAD
MOV       1 D00004	// 상태_방향 0없음 1상승 2하강
MPOP
AND       M00006	// 판단_아래요청 판단층보다 아래에 요청 있음
LOAD<>    D00004 1	// 상태_방향 0없음 1상승 2하강
OR NOT    M00005	// 판단_위요청 판단층보다 위에 요청 있음
AND LOAD
MOV       2 D00004	// 상태_방향 0없음 1상승 2하강
// output comment: 위요청이 있고 아래요청이 없을 때 상승방향 위요청이 있고 아래요청이 있으면(내려가는 경우가 아니라고 할 때) 상승방향 유지  
// 도착상태에서 대기, 상승, 하강상태중 하나로 전이
; L24
LOAD=     D00010 3	// 상태_운행 0대기 1상승 2하강 3도착 8점검 9에러
AND       M00004	// 문_동작완료 닫힘 4초 + 문닫힘
MPUSH
AND=      D00004 0	// 상태_방향 0없음 1상승 2하강
MOV       0 D00010	// 상태_운행 0대기 1상승 2하강 3도착 8점검 9에러
MLOAD
AND=      D00004 1	// 상태_방향 0없음 1상승 2하강
MOV       1 D00010	// 상태_운행 0대기 1상승 2하강 3도착 8점검 9에러
MPOP
AND=      D00004 2	// 상태_방향 0없음 1상승 2하강
MOV       2 D00010	// 상태_운행 0대기 1상승 2하강 3도착 8점검 9에러

PROGRAM P08_OUPUT (task: 스캔 프로그램)

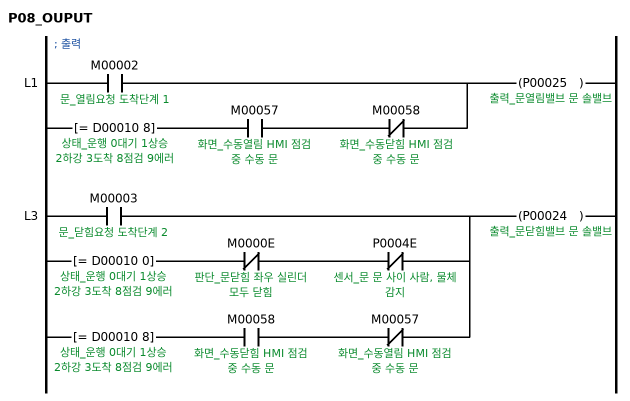
// 출력
; L1
LOAD      M00002	// 문_열림요청 도착단계 1
LOAD=     D00010 8	// 상태_운행 0대기 1상승 2하강 3도착 8점검 9에러
AND       M00057	// 화면_수동열림 HMI 점검 중 수동 문
AND NOT   M00058	// 화면_수동닫힘 HMI 점검 중 수동 문
OR LOAD
OUT       P00025	// 출력_문열림밸브 문 솔밸브
; L3
LOAD      M00003	// 문_닫힘요청 도착단계 2
LOAD=     D00010 0	// 상태_운행 0대기 1상승 2하강 3도착 8점검 9에러
AND NOT   M0000E	// 판단_문닫힘 좌우 실린더 모두 닫힘
AND NOT   P0004E	// 센서_문 문 사이 사람, 물체 감지
OR LOAD
LOAD=     D00010 8	// 상태_운행 0대기 1상승 2하강 3도착 8점검 9에러
AND       M00058	// 화면_수동닫힘 HMI 점검 중 수동 문
AND NOT   M00057	// 화면_수동열림 HMI 점검 중 수동 문
OR LOAD
OUT       P00024	// 출력_문닫힘밸브 문 솔밸브

PROGRAM INIT (task: INIT)

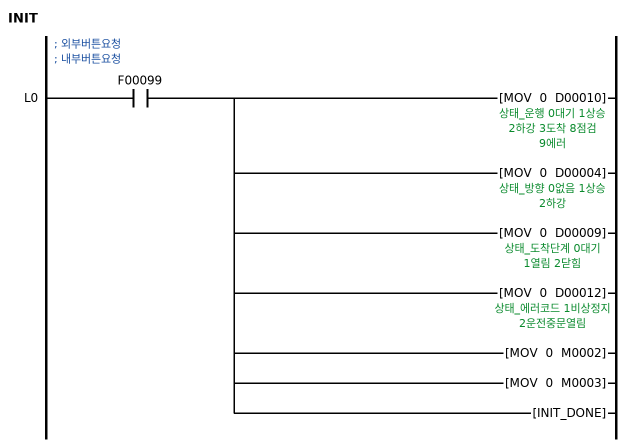
; L0
LOAD      F00099
MOV       0 D00010	// 상태_운행 0대기 1상승 2하강 3도착 8점검 9에러
MOV       0 D00004	// 상태_방향 0없음 1상승 2하강
MOV       0 D00009	// 상태_도착단계 0대기 1열림 2닫힘
MOV       0 D00012	// 상태_에러코드 1비상정지 2운전중문열림
MOV       0 M0002
MOV       0 M0003
INIT_DONE
// output comment: 외부버튼요청
// output comment: 내부버튼요청

VARIABLES AND COMMENTS (devices not used above)
P0004C	BIT	센서_우문열림 // 문 실린더 센서
P0004A	BIT	센서_좌문열림 // 문 실린더 센서